Universal Robots URScript: T011_codellama_34b_baseline_rep1_retry2.urscript

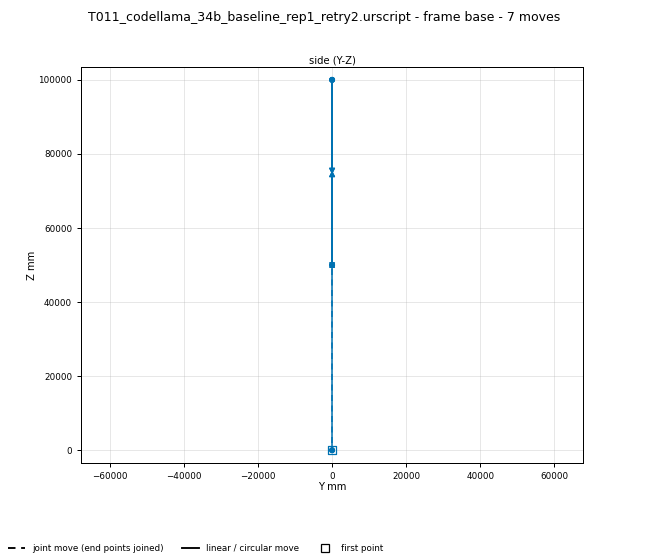
[picture p0: tool path of T011_codellama_34b_baseline_rep1_retry2.urscript in frame base, 7 of 7 moves have a stored position in this frame; points joined in program order, loops and branches not executed]
def dual_zone_pick_place():
    # Home the robot arm
    movej(p[0, 0, 0, 0, 0, 0], v=250.0)

    # Move above storage bin
    movel(p[0, 0, 100, 0, 0, 0], v=280.0)

    # Descend to pick
    movel(p[0, 0, 50, 0, 0, 0], v=120.0)

    # Lift from bin
    movel(p[0, 0, 100, 0, 0, 0], v=200.0)

    # Transit to handoff zone
    movel(p[0, 0, 50, 0, 0, 0], v=250.0)

    # Place in handoff zone
    movej(p[0, 0, 100, 0, 0, 0], v=250.0)

    # Return to home position
    movej(p[0, 0, 0, 0, 0, 0], v=250.0)
